(* IEC 61131-3 sources: Pirate/PLC/DUT, 7 files *)

(* ---- ST_AreteZone.st ---- *)
TYPE ST_AreteZone :
STRUCT
    NoeudA : UINT; // indice dans le tableau des noeuds de la zone
    NoeudB : UINT; // indice dans le tableau des noeuds de la zone
    EquipementIndex : INT; // -1 pour une liaison permanente, sinon indice equipement
END_STRUCT
END_TYPE

(* ---- ST_ConnexionPorts.st ---- *)
TYPE ST_ConnexionPorts :
STRUCT
    Id : UINT;
    PosteA : UINT;
    PortA : UINT;
    PosteB : UINT;
    PortB : UINT;
END_STRUCT
END_TYPE

(* ---- ST_Equipement.st ---- *)
TYPE ST_Equipement :
STRUCT
    Id : UINT; // identifiant local au poste
    NoeudA : UINT; // noeud local
    NoeudB : UINT; // noeud local
    Ferme : BOOL;
    Defaut : BOOL;
    Conducteur : BOOL; // calcule, ne pas commander
END_STRUCT
END_TYPE

(* ---- ST_Noeud.st ---- *)
TYPE ST_Noeud :
STRUCT
    IdLocal : UINT;
    IdZone : UINT; // affecte par FB_Zone
    SousTension : BOOL; // resultat BFS
END_STRUCT
END_TYPE

(* ---- ST_Port.st ---- *)
TYPE ST_Port :
STRUCT
    Id : UINT;
    NoeudLocal : UINT; // plusieurs connexions externes autorisees
END_STRUCT
END_TYPE

(* ---- ST_RefNoeud.st ---- *)
TYPE ST_RefNoeud :
STRUCT
    PosteId : UINT;
    NoeudLocal : UINT;
    NoeudZone : UINT;
END_STRUCT
END_TYPE

(* ---- ST_Source.st ---- *)
TYPE ST_Source :
STRUCT
    Id : UINT;
    NoeudLocal : UINT; // noeud interne a la sous-station
    Active : BOOL;
END_STRUCT
END_TYPE
